(* IEC 61131-3 sources: Caravan/Archiv/12-04-19/Stations/Terminal/HMI/Network/NewAgeAlarmVis, 1 file *)

(* ---- ONE_NewAgeAlarmVis_Table.st ---- *)
#define OBJECTS_CONFIG

#include "..\..\Class\AlarmDisplayList\AlarmTemp.h"
//Define part of class TitleLine
// Eigenschaften des UDCs
//----------------------------------------------------------------------------------------------------------------------------
#define   TitleLine_UDCVersion                2           // Version des aktuellen UDCs (sprdie v1.2 changed from 1 -> 2)
#define   TitleLine_VariableNo                8           // Anzahl der Variablen, die dem UDC mitgegeben werden (sprdie v1.2 changed from 6 -> 8)
#define   TitleLine_BoolNo                    1           // Anzahl der Boolschen-Variablen, die dem UDC mitgegeben werden
#define   TitleLine_TextschemeNo              1           // Anzahl der Textschemen, die dem UDC mitgegeben werden
#include "..\..\Class\AlarmTitleLine\Alarms.h"

FUNCTION GLOBAL TAB ONE_NewAgeAlarmVis
-1$UINT, 0$UINT,
1$UINT, 0$UINT,

11$UDINT,
TO_UDINT(1738954212), "_AlarmDisplay", 0$UINT, 10$UINT, 0$UINT,
TO_UDINT(3745297859), "_Bit32", 0$UINT, 1$UINT, 1$UINT,
TO_UDINT(2980745877), "_MyIO", 0$UINT, 3$UINT, 0$UINT,
TO_UDINT(3043040051), "_ScrollArea", 0$UINT, 15$UINT, 0$UINT,
TO_UDINT(3279795640), "AlarmDisplayList", 1$UINT, 7$UINT, 1$UINT,
TO_UDINT(718326546), "AlarmTitleLine", 1$UINT, 1$UINT, 1$UINT,
TO_UDINT(2225119864), "MerkerEx", 1$UINT, 21$UINT, 2$UINT,
TO_UDINT(1850111279), "String", 1$UINT, 10$UINT, 2$UINT,
TO_UDINT(2898603620), "StringInternal", 1$UINT, 82$UINT, 0$UINT,
TO_UDINT(112430022), "TitleLine", 1$UINT, 3$UINT, 0$UINT,
TO_UDINT(3232495061), "VirtualBaseInit", 1$UINT, 3$UINT, 0$UINT,

_NO_ATTR, TO_UDINT(2843603871), "_BITALARMTITLE",

_NO_ATTR, TO_UDINT(3279795640), "ALARMDISPLAYLIST",

_NO_ATTR, TO_UDINT(1387240034), "ALARMTITLE",

1$UINT, TO_UDINT(3116160222), "ALARMDISPLAYLIST\ALARMTXTLONG\MERKEREX0",
1$UINT, TO_UDINT(2022897073), "ALARMDISPLAYLIST\ALARMTXTSHORT\MERKEREX0",

1$UINT, TO_UDINT(358957295), "ALARMDISPLAYLIST\ALARMTXTLONG",
1$UINT, TO_UDINT(3350483968), "ALARMDISPLAYLIST\ALARMTXTSHORT",

//Internal connections
0$UDINT,
4$UDINT,
TO_UDINT(1), "AlarmTxtShort", TO_UDINT(6),
TO_UDINT(1), "AlarmTxtLong", TO_UDINT(5),
TO_UDINT(5), "MerkerEx0", TO_UDINT(3),
TO_UDINT(6), "MerkerEx0", TO_UDINT(4),
0$UDINT,
5$UDINT,
TO_UDINT(1), "ColumnChoice", TO_UDINT(0), "Data",
TO_UDINT(1), "coAlarmTitle", TO_UDINT(2), "Server0",
TO_UDINT(2), "ColumnChoice", TO_UDINT(0), "Data",
TO_UDINT(5), "DataBuffer", TO_UDINT(3), "m_udLength",
TO_UDINT(6), "DataBuffer", TO_UDINT(4), "m_udLength",

//Initialization values
0$UDINT,
12$UDINT,
TO_UDINT(0), "", TO_UDINT(2#11101),//|NewAgeAlarmVis._BitAlarmTitle.Data;
TO_UDINT(1), "VerticalLevel", TO_UDINT(1),//|NewAgeAlarmVis.AlarmDisplayList.VerticalLevel;
TO_UDINT(1), "LineWidth", TO_UDINT(10000),//|NewAgeAlarmVis.AlarmDisplayList.LineWidth;
TO_UDINT(1), "ExtendedScrollBar", TO_UDINT(1),//|NewAgeAlarmVis.AlarmDisplayList.ExtendedScrollBar;
TO_UDINT(1), "HistoryTemporary", TO_UDINT(1),//|NewAgeAlarmVis.AlarmDisplayList.HistoryTemporary;
TO_UDINT(1), "MaxNo", TO_UDINT(100),//|NewAgeAlarmVis.AlarmDisplayList.MaxNo;
TO_UDINT(1), "Filter", TO_UDINT(2#01101),//|NewAgeAlarmVis.AlarmDisplayList.Filter;
TO_UDINT(1), "coAlarmTitle", TO_UDINT(0),//|NewAgeAlarmVis.AlarmDisplayList.coAlarmTitle;
TO_UDINT(3), "ThreadSafe", TO_UDINT(0),//|NewAgeAlarmVis.AlarmTxtLong\AlarmDisplayList\MerkerEx0.ThreadSafe;
TO_UDINT(4), "ThreadSafe", TO_UDINT(0),//|NewAgeAlarmVis.AlarmTxtShort\AlarmDisplayList\MerkerEx0.ThreadSafe;
TO_UDINT(5), "SingleRealloc", TO_UDINT(1),//|NewAgeAlarmVis.AlarmDisplayList\AlarmTxtLong.SingleRealloc;
TO_UDINT(6), "SingleRealloc", TO_UDINT(1),//|NewAgeAlarmVis.AlarmDisplayList\AlarmTxtShort.SingleRealloc;

//Symbolic initialization values
0$UDINT,
0$UDINT,

//Initialization of string values
0$UDINT,
0$UDINT,

//Configuration of tasks (RealTime, Cyclic, Background)
0$UDINT,
0$UDINT,

0$UDINT,
0$UDINT,

0$UDINT,
0$UDINT,

//External connections
0$UDINT,
4$UDINT,
TO_UDINT(1), "Lse", C_DIR, TO_UDINT(299963966), "Lse","Lse",
TO_UDINT(1), "coSystemLogging", C_TRY, TO_UDINT(2516821708), "SystemLogging1","ClassSvr",
TO_UDINT(2), "Lse", C_DIR, TO_UDINT(299963966), "Lse","Lse",
TO_UDINT(2), "coSystemLogging", C_TRY, TO_UDINT(2516821708), "SystemLogging1","ClassSvr",

//Magic internal connections
0$UDINT,
0$UDINT,

//Configuration of timeslots of tasks (RealTime, Cyclic)
#ifdef __LSLLDR_TIMESLOTS__
0$UDINT,
0$UDINT,

0$UDINT,
0$UDINT,

#endif //__LSLLDR_TIMESLOTS__

//MultiMaster connections
#ifdef __LSLLDR_MULTIMASTER__
0$UDINT,
0$UDINT,
#endif //__LSLLDR_MULTIMASTER__

//Configuration for task ID (RealTime, CyclicTime)
#ifdef __LSLLDR_TASKID__
"\\\\TASKS2  "
0$UDINT,
0$UDINT,

0$UDINT,
0$UDINT,

0$UDINT,
0$UDINT,

#endif //__LSLLDR_TASKID__

END_FUNCTION
